Staubli VAL3: init.pgx

program init()
begin
  //应用初始化：可重复调用（幂等）
  nState=0
  nAlarm=0
  sAlarmMsg=""
  bStartCmd=false
  bStopCmd=false
  bPauseCmd=false
  bResetCmd=false
  bRunning=false
  nCycleCount=0
  nProdCount=0
end
